Yaskawa INFORM job: OBLICZ_SZLIF_TROJNIKA.JBI

/JOB
//NAME OBLICZ_SZLIF_TROJNIKA
///FOLDERNAME TROJNIKI
//POS
///NPOS 0,0,0,4,0,0
///USER 10
///TOOL 17
///POSTYPE USER
///RECTAN
///RCONF 1,0,0,0,0,0,0,0,0,0,0,0,0,0,0,0,0,0,0,0,0,0,0,0
P00010=63.000,1.000,-2.000,-90.0000,-90.0000,90.0000
///USER 8
P00011=8.000,1.000,-2.000,-90.0000,-90.0000,90.0000
P00012=63.000,1.000,10.000,-90.0000,-90.0000,90.0000
///RCONF 0,0,0,0,0,0,0,0,0,0,0,0,0,0,0,0,0,0,0,0,0,0,0,0
P00013=8.000,1.000,10.000,-90.0000,-90.0000,90.0000
//INST
///DATE 2026/11/18 08:00
///ATTR SC,RW
///GROUP1 RB1
NOP
'FREZ 12MM TOOL 17
'START OSI FREZA: PROMIEN 3MM
'I073: KROK SREDNICY W 0.001MM
'D120: PROMIEN DOCELOWY
'D121: KROK PROMIENIA NA SZTUKE
'D103-D105 Z TROJNIK_TEST
*PARAMETRY
IFTHENEXP I035=30
	 NOP
ELSE
	 PAUSE
	 JUMP *PARAMETRY
ENDIF
IFTHENEXP I120<1
	 PAUSE
	 JUMP *PARAMETRY
ENDIF
IFTHENEXP I120=1
	'NOWA SZTUKA: SREDNICE
	 IFTHENEXP I070<=0
		 PAUSE
		 JUMP *PARAMETRY
	 ENDIF
	 IFTHENEXP I074<0
		 PAUSE
		 JUMP *PARAMETRY
	 ENDIF
	 SET D073  EXPRESS I071 * 100
	 SET D075  EXPRESS I074 * 100
	 MUL D075 2
	 SET D072  EXPRESS I070 * 100
	 SET D079 D072
	 SET D120  EXPRESS D073 - D075 - D072
	 DIV D120 2
	 IFTHENEXP D120<3000
		 PAUSE
		 JUMP *PARAMETRY
	 ENDIF
	'KROK SREDNICY: DODATNI PARZYSTY
	 SET D121 I073
	 IFTHENEXP D121<2
		 PAUSE
		 JUMP *PARAMETRY
	 ENDIF
	 SET D066 D121
	 DIV D066 2
	 MUL D066 2
	 IFTHENEXP D066=D121
		 DIV D121 2
	 ELSE
		 PAUSE
		 JUMP *PARAMETRY
	 ENDIF
	 SET B030 0
	 DOUT OT#(6) OFF
	 SET D089  EXPRESS I089 * 1000
ELSE
	 IFTHENEXP D121<=0
		 PAUSE
		 JUMP *PARAMETRY
	 ENDIF
	 IFTHENEXP D120<3000
		 PAUSE
		 JUMP *PARAMETRY
	 ENDIF
ENDIF
'PROMIEN Z NUMERU OBIEGU
SET D074  EXPRESS I120 - 1
MUL D074 D121
ADD D074 3000
'OSTATNI KROK DO GRANICY
IFTHENEXP D074>D120
	 SET D074 D120
ENDIF
'PUNKTY DLA TOOL 17
FOR I060 START= 10 TO 13 STEP= 1
	 SETE P[I060] TL#(17)
NEXT I060
'TABELA PARAMETROW DLA SREDNIC
'D032-D035: Offset Start Z (Dol,
'Gora, Prawy, Lewy)
''''''''''''''''''
SWITCH I035
CASE 30
	''''''''
	'26,9mm'
	''''''''
	'wysokosc spawu'
	'gora dol'
	 SET D032 19000
	'gora
	 SET D033 0
	'prawo
	 SET D034 0
	'dol
	 SET D035 0
	'ustawienia katow
	 SET D069 -1800000
	 SET D070 0
	 SET D071 900000
	 SETE P010 (4) D069
	 SETE P010 (5) D070
	 SETE P010 (6) D071
	 SETE P011 (4) D069
	 SETE P011 (5) D070
	 SETE P011 (6) D071
	 SETE P012 (4) D069
	 SETE P012 (5) D070
	 SETE P012 (6) D071
	 SETE P013 (4) D069
	 SETE P013 (5) D070
	 SETE P013 (6) D071
ENDSWITCH
'''''''''''''''''''''
'pozycja szlifowania'
''''''''lewo'''''''''
'''''''''''''''''''''
SET D066  EXPRESS 0 + D103 + D074
SET D067  EXPRESS 0 + D104
SET D068  EXPRESS D032 + D105
SETE P010 (1) D066
SETE P010 (2) D067
SETE P010 (3) D068
'''''''''''''''''''''
'pozycja szlifowania'
''''''''gora'''''''''
'''''''''''''''''''''
SET D066  EXPRESS 0 + D103
SET D067  EXPRESS 0 + D104 - D074
SETE P011 (1) D066
SETE P011 (2) D067
SETE P011 (3) D068
'''''''''''''''''''''
'pozycja szlifowania'
''''''''prawo''''''''
'''''''''''''''''''''
SET D066  EXPRESS 0 + D103 - D074
SET D067  EXPRESS 0 + D104
SETE P012 (1) D066
SETE P012 (2) D067
SETE P012 (3) D068
'''''''''''''''''''''
'pozycja szlifowania'
'''''''''dol'''''''''
'''''''''''''''''''''
SET D066  EXPRESS 0 + D103
SET D067  EXPRESS 0 + D104 + D074
SETE P013 (1) D066
SETE P013 (2) D067
SETE P013 (3) D068
RET
END
